RoboDK station: PickAndPlace.rdk

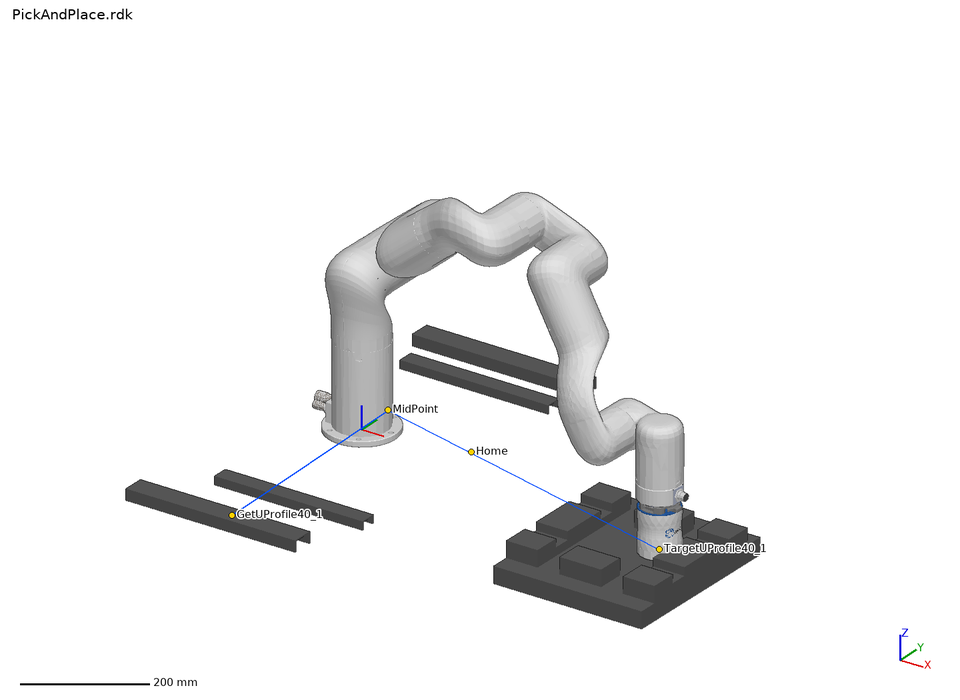
[picture v0: the station drawn from its stored meshes, robots at their saved joint values, targets as dots, program paths as lines]
Station PickAndPlace (saved by RoboDK 6.2.0). Poses are relative to the parent item; angles as X-Y-Z fixed-axis rotations.
  - frame uFactory xArm6 Base at (-50, 0, 100) mm
    - robot uFactory xArm6: 6 axes, payload 5 kg, reach 700 mm, repeatability 0.1 mm, weight 12.2 kg
        modified DH rows (alpha deg, a mm, theta deg, d mm): 0, 0, 0, 267; -90, 0, -79.35, 0; 0, 289.489, 79.35, 0; -90, 77.5, 0, 342.5; 90, 0, 0, 0; -90, 76, 0, 97
        joint limits [-360, -118, -225, -360, -97, -360] to [360, 120, 11, 360, 180, 360]; home [0, 0, 0, 0, 0, 0]; saved at [0.172, 51.288, -79.25, 0, 27.962, 92.672]
      - tool OnRobot MG10 Magnetic Gripper, TCP at (0, 0, 90) mm, size 71 x 74.9 x 91.4 mm
    - target Home (Cartesian target) at (207, 0, 19) mm, rotated rx -180 ry 0 rz 0 deg; joints [0, 0, 0, 0, 0, 0] of uFactory xArm6
    - target GetUProfile40_1 (Cartesian target) at (9.13, -363.2, 0) mm, rotated rx -180 ry 0 rz -11 deg; joints [-88.559, 20.873, -30.902, 0.002, 10.029, -77.562] of uFactory xArm6
    - target MidPoint (Cartesian target) at (231.62, -260.08, 201.95) mm, rotated rx 179.56 ry 1.61 rz 20.91 deg; joints [-47.71, -18.36, -31.47, -2.17, 50.03, -67.23] of uFactory xArm6
    - target TargetUProfile40_1 (Cartesian target) at (560.5, 1.68, -50) mm, rotated rx 180 ry 0 rz -92.5 deg; joints [0.172, 51.288, -79.25, 0, 27.962, 92.672] of uFactory xArm6
  - object Mask at (450, 0, 0) mm, rotated rx 90 ry 0 rz 90 deg, size 320 x 60 x 280 mm, geometry from Mask.step
  - object UProfile30_1 at (0, -250, 100) mm, rotated rx -90 ry 0 rz 0 deg, size 280 x 15 x 30 mm, geometry from UProfile30.step
  - object UProfile30_2 at (0, 250, 100) mm, rotated rx -90 ry 0 rz 0 deg, size 280 x 15 x 30 mm, geometry from UProfile30.step
  - object UProfile40_1 at (0, -350, 100) mm, rotated rx -90 ry 0 rz 0 deg, size 320 x 20 x 40 mm, geometry from UProfile40.step
  - object UProfile40_2 at (50, 350, 100) mm, rotated rx -90 ry 0 rz 0 deg, size 320 x 20 x 40 mm, geometry from UProfile40.step
  - program Home (3 instructions, listed below)
  - program PickAndPlaceUProfile40_1 (7 instructions, listed below)
  - program Main (3 instructions, listed below)
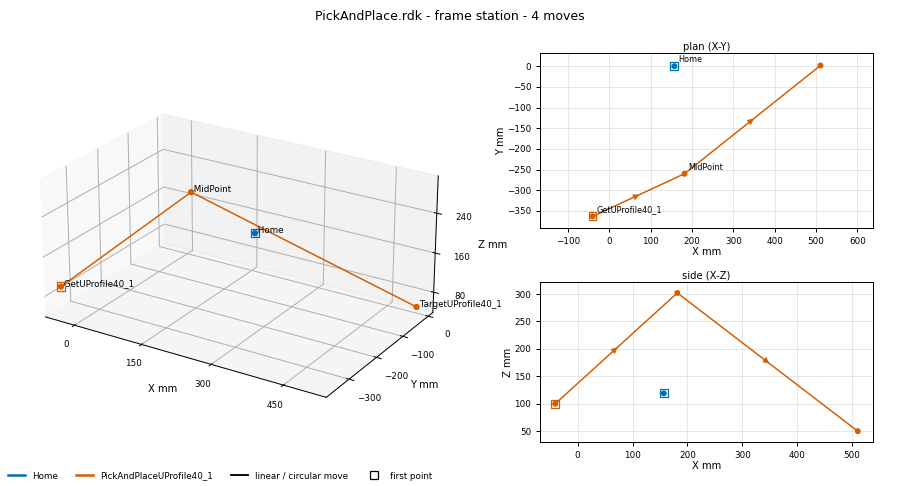
[picture p0: tool path of PickAndPlace.rdk in frame station, 4 of 4 moves have a stored position in this frame; points joined in program order, loops and branches not executed]

--- program Home (robot uFactory xArm6) ---
  Set Ref.: uFactory xArm6 Base
  Set Tool: OnRobot MG10 Magnetic Gripper
  MoveJ (Home)

--- program PickAndPlaceUProfile40_1 (robot uFactory xArm6) ---
  Set Ref.: uFactory xArm6 Base
  Set Tool: OnRobot MG10 Magnetic Gripper
  MoveJ (GetUProfile40_1)
  Attach to OnRobot MG10 Magnetic Gripper
  MoveL (MidPoint)
  MoveL (TargetUProfile40_1)
  Detach from OnRobot MG10 Magnetic Gripper

--- program Main (robot uFactory xArm6) ---
  Call Home
  Call PickAndPlaceUProfile40_1
  Call Home
